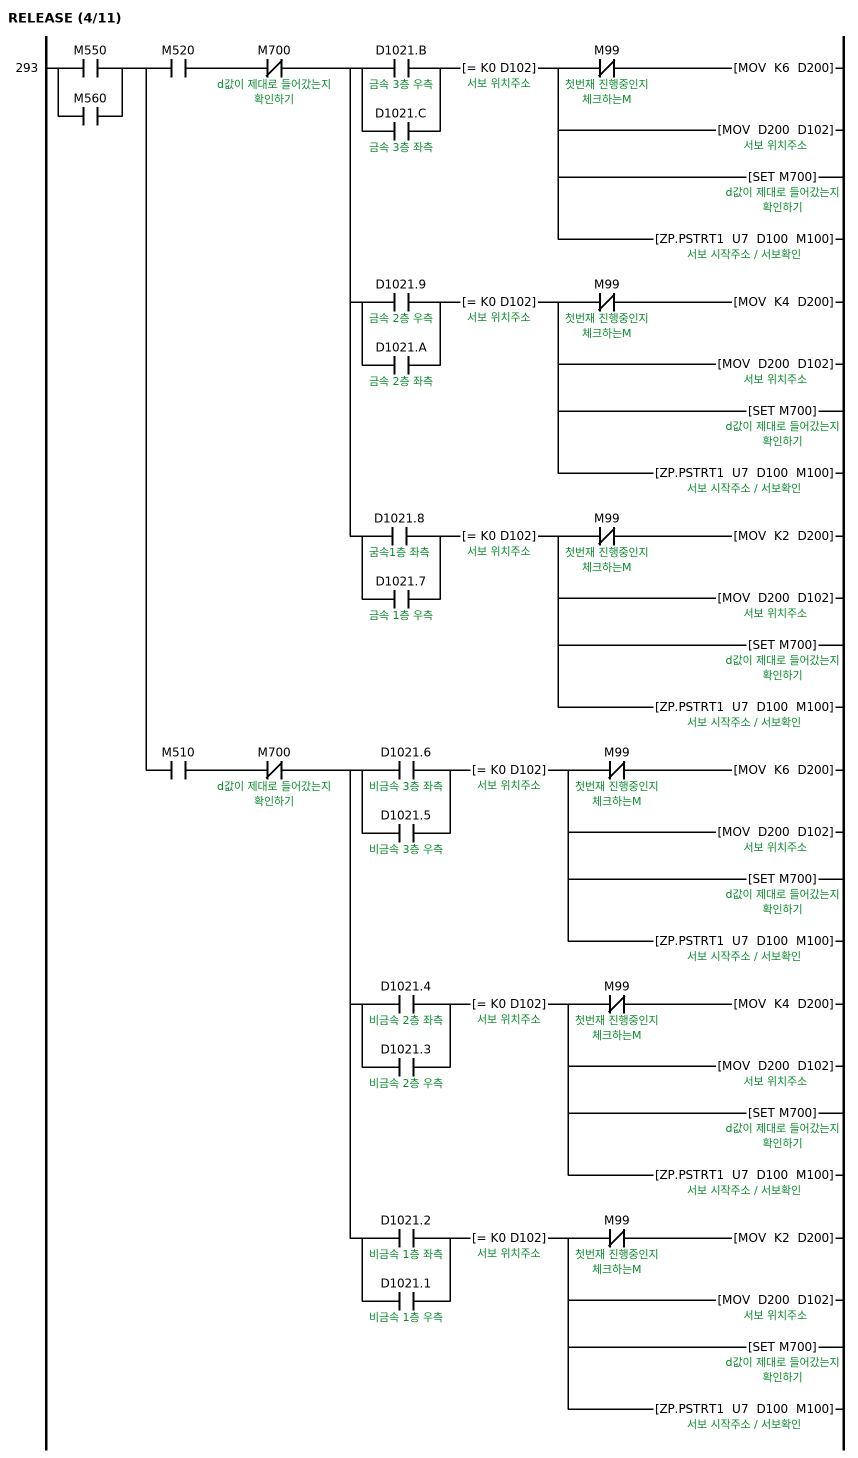
[picture p24: ladder of RELEASE, rungs at steps 293 to 293]
293   LD      M550
      OR      M560
      MPS
      AND     M520
      ANI     M700  ; d값이 제대로 들어갔는지 확인하기
      MPS
      LD      D1021.B  ; 금속 3층 우측
      OR      D1021.C  ; 금속 3층 좌측
      ANB
      AND=    K0 D102  ; 서보 위치주소
      MPS
      ANI     M99  ; 첫번재 진행중인지 체크하는M
      MOV     K6 D200
      MPP
      MOV     D200 D102
      SET     M700  ; d값이 제대로 들어갔는지 확인하기
      ZP.PSTRT1 U7 D100 M100  ; 서보 시작주소 / 서보확인
      MRD
      LD      D1021.9  ; 금속 2층 우측
      OR      D1021.A  ; 금속 2층 좌측
      ANB
      AND=    K0 D102  ; 서보 위치주소
      MPS
      ANI     M99  ; 첫번재 진행중인지 체크하는M
      MOV     K4 D200
      MPP
      MOV     D200 D102
      SET     M700  ; d값이 제대로 들어갔는지 확인하기
      ZP.PSTRT1 U7 D100 M100
      MPP
      LD      D1021.8  ; 굼속1층 좌측
      OR      D1021.7  ; 금속 1층 우측
      ANB
      AND=    K0 D102  ; 서보 위치주소
      MPS
      ANI     M99  ; 첫번재 진행중인지 체크하는M
      MOV     K2 D200
      MPP
      MOV     D200 D102
      SET     M700  ; d값이 제대로 들어갔는지 확인하기
      ZP.PSTRT1 U7 D100 M100
      MPP
      AND     M510
      ANI     M700  ; d값이 제대로 들어갔는지 확인하기
      MPS
      LD      D1021.6  ; 비금속 3층 좌측
      OR      D1021.5  ; 비금속 3층 우측
      ANB
      AND=    K0 D102  ; 서보 위치주소
      MPS
      ANI     M99  ; 첫번재 진행중인지 체크하는M
      MOV     K6 D200
      MPP
      MOV     D200 D102
      SET     M700  ; d값이 제대로 들어갔는지 확인하기
      ZP.PSTRT1 U7 D100 M100
      MRD
      LD      D1021.4  ; 비금속 2층 좌측
      OR      D1021.3  ; 비금속 2층 우측
      ANB
      AND=    K0 D102  ; 서보 위치주소
      MPS
      ANI     M99  ; 첫번재 진행중인지 체크하는M
      MOV     K4 D200
      MPP
      MOV     D200 D102
      SET     M700  ; d값이 제대로 들어갔는지 확인하기
      ZP.PSTRT1 U7 D100 M100
      MPP
      LD      D1021.2  ; 비금속 1층 좌측
      OR      D1021.1  ; 비금속 1층 우측
      ANB
      AND=    K0 D102  ; 서보 위치주소
      MPS
      ANI     M99  ; 첫번재 진행중인지 체크하는M
      MOV     K2 D200
      MPP
      MOV     D200 D102
      SET     M700  ; d값이 제대로 들어갔는지 확인하기
      ZP.PSTRT1 U7 D100 M100
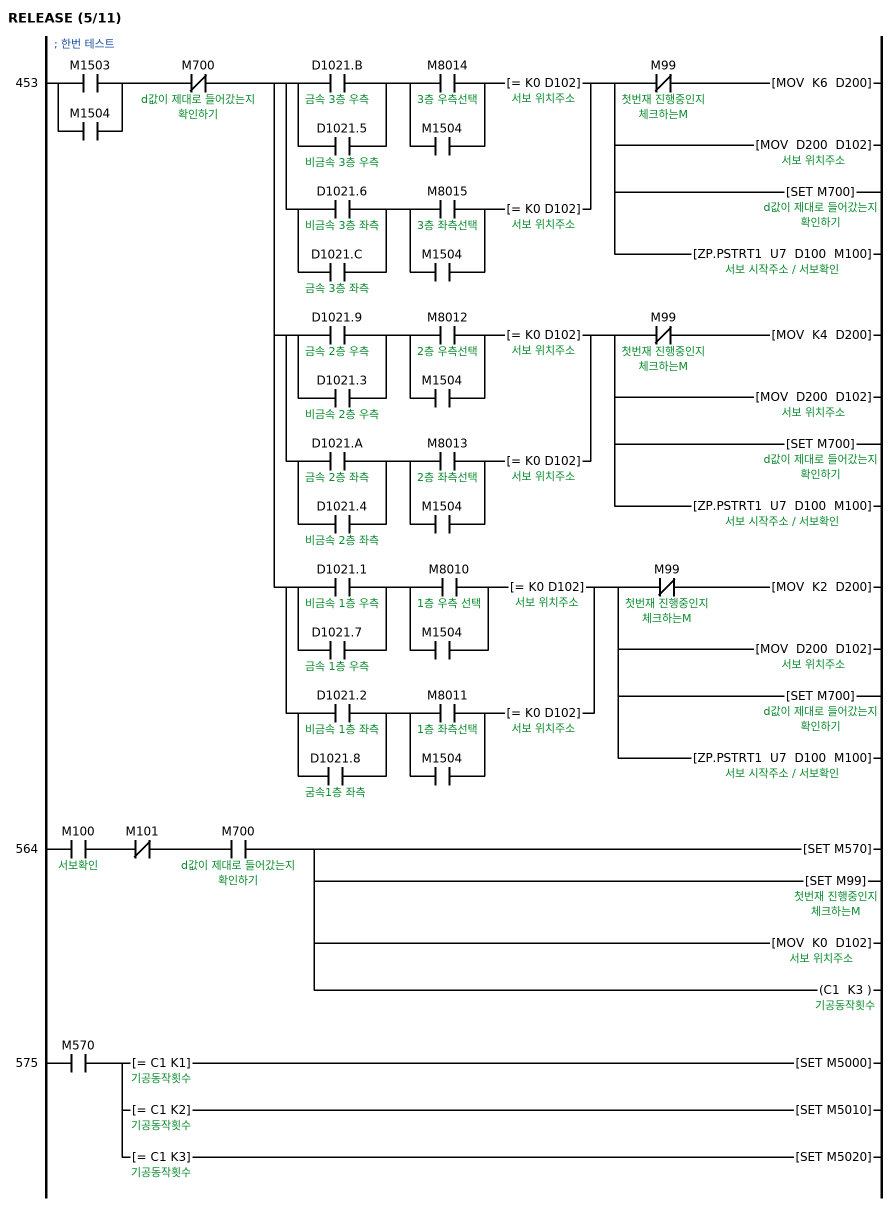
; 한번 테스트
453   LD      M1503
      OR      M1504
      ANI     M700  ; d값이 제대로 들어갔는지 확인하기
      MPS
      LD      D1021.B  ; 금속 3층 우측
      OR      D1021.5  ; 비금속 3층 우측
      LD      M8014  ; 3층 우측선택
      OR      M1504
      ANB
      AND=    K0 D102  ; 서보 위치주소
      LD      D1021.6  ; 비금속 3층 좌측
      OR      D1021.C  ; 금속 3층 좌측
      LD      M8015  ; 3층 좌측선택
      OR      M1504
      ANB
      AND=    K0 D102  ; 서보 위치주소
      ORB
      ANB
      MPS
      ANI     M99  ; 첫번재 진행중인지 체크하는M
      MOV     K6 D200
      MPP
      MOV     D200 D102
      SET     M700  ; d값이 제대로 들어갔는지 확인하기
      ZP.PSTRT1 U7 D100 M100
      MRD
      LD      D1021.9  ; 금속 2층 우측
      OR      D1021.3  ; 비금속 2층 우측
      LD      M8012  ; 2층 우측선택
      OR      M1504
      ANB
      AND=    K0 D102  ; 서보 위치주소
      LD      D1021.A  ; 금속 2층 좌측
      OR      D1021.4  ; 비금속 2층 좌측
      LD      M8013  ; 2층 좌측선택
      OR      M1504
      ANB
      AND=    K0 D102  ; 서보 위치주소
      ORB
      ANB
      MPS
      ANI     M99  ; 첫번재 진행중인지 체크하는M
      MOV     K4 D200
      MPP
      MOV     D200 D102
      SET     M700  ; d값이 제대로 들어갔는지 확인하기
      ZP.PSTRT1 U7 D100 M100
      MPP
      LD      D1021.1  ; 비금속 1층 우측
      OR      D1021.7  ; 금속 1층 우측
      LD      M8010  ; 1층 우측 선택
      OR      M1504
      ANB
      AND=    K0 D102  ; 서보 위치주소
      LD      D1021.2  ; 비금속 1층 좌측
      OR      D1021.8  ; 굼속1층 좌측
      LD      M8011  ; 1층 좌측선택
      OR      M1504
      ANB
      AND=    K0 D102  ; 서보 위치주소
      ORB
      ANB
      MPS
      ANI     M99  ; 첫번재 진행중인지 체크하는M
      MOV     K2 D200
      MPP
      MOV     D200 D102
      SET     M700  ; d값이 제대로 들어갔는지 확인하기
      ZP.PSTRT1 U7 D100 M100
564   LD      M100  ; 서보확인
      ANI     M101
      AND     M700  ; d값이 제대로 들어갔는지 확인하기
      SET     M570
      SET     M99  ; 첫번재 진행중인지 체크하는M
      MOV     K0 D102
      OUT     C1 K3  ; 기공동작횟수
575   LD      M570
      MPS
      AND=    C1 K1  ; 기공동작횟수
      SET     M5000
      MRD
      AND=    C1 K2  ; 기공동작횟수
      SET     M5010
      MPP
      AND=    C1 K3  ; 기공동작횟수
      SET     M5020
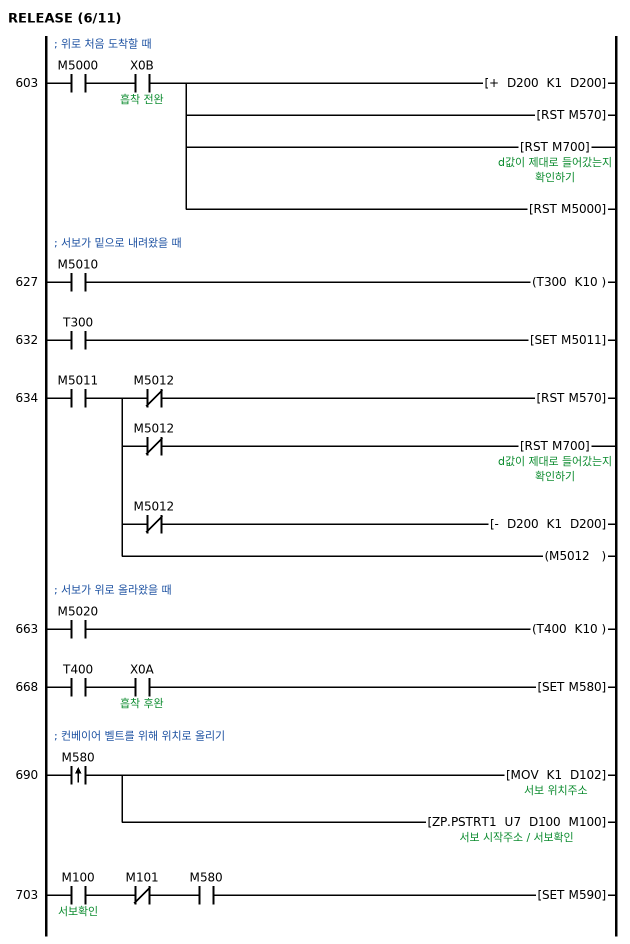
; 위로 처음 도착할 때
603   LD      M5000
      AND     X0B  ; 흡착 전완
      +       D200 K1 D200
      RST     M570
      RST     M700  ; d값이 제대로 들어갔는지 확인하기
      RST     M5000
; 서보가 밑으로 내려왔을 때
627   LD      M5010
      OUT     T300 K10
632   LD      T300
      SET     M5011
634   LD      M5011
      MPS
      ANI     M5012
      RST     M570
      MRD
      ANI     M5012
      RST     M700  ; d값이 제대로 들어갔는지 확인하기
      MRD
      ANI     M5012
      -       D200 K1 D200
      MPP
      OUT     M5012
; 서보가 위로 올라왔을 때
663   LD      M5020
      OUT     T400 K10
668   LD      T400
      AND     X0A  ; 흡착 후완
      SET     M580
; 컨베이어 벨트를 위해 위치로 올리기
690   LDP     M580
      MOV     K1 D102
      ZP.PSTRT1 U7 D100 M100
703   LD      M100  ; 서보확인
      ANI     M101
      AND     M580
      SET     M590
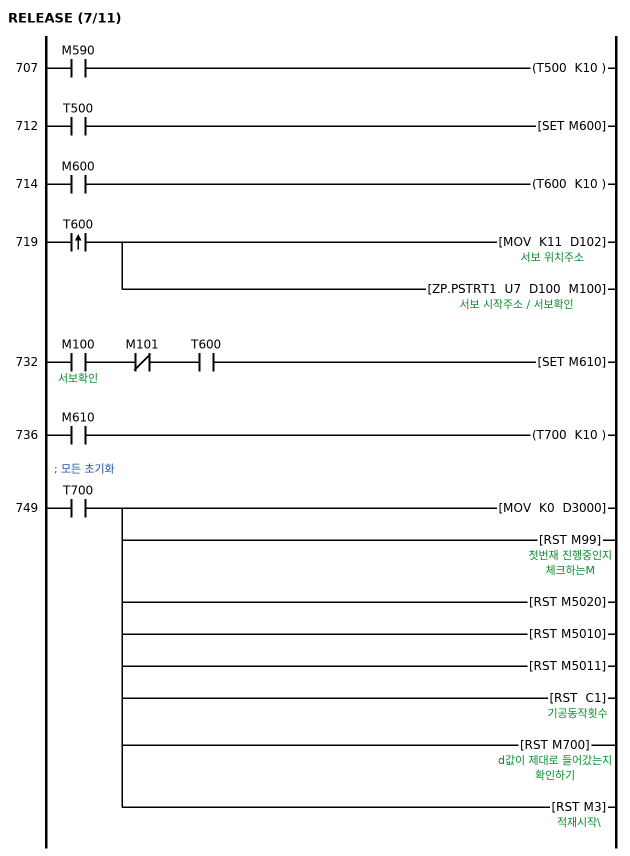
707   LD      M590
      OUT     T500 K10
712   LD      T500
      SET     M600
714   LD      M600
      OUT     T600 K10
719   LDP     T600
      MOV     K11 D102
      ZP.PSTRT1 U7 D100 M100
732   LD      M100  ; 서보확인
      ANI     M101
      AND     T600
      SET     M610
736   LD      M610
      OUT     T700 K10
; 모든 초기화
749   LD      T700
      MOV     K0 D3000
      RST     M99  ; 첫번재 진행중인지 체크하는M
      RST     M5020
      RST     M5010
      RST     M5011
      RST     C1  ; 기공동작횟수
      RST     M700  ; d값이 제대로 들어갔는지 확인하기
      RST     M3  ; 적재시작\
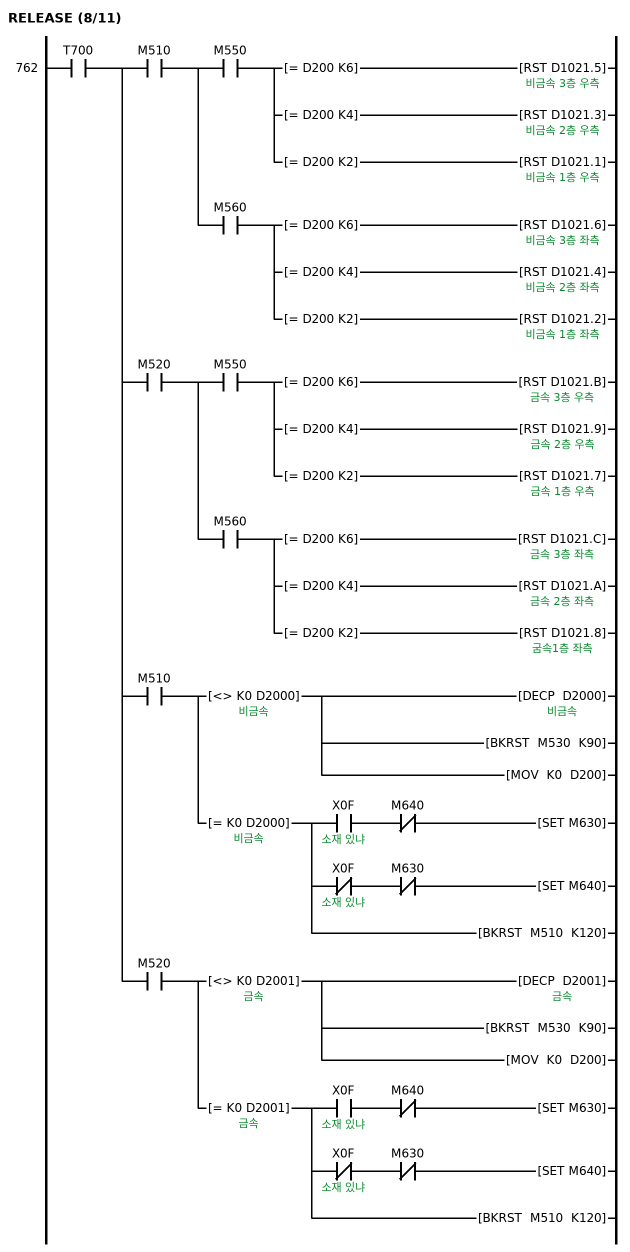
762   LD      T700
      MPS
      AND     M510
      MPS
      AND     M550
      MPS
      AND=    D200 K6
      RST     D1021.5  ; 비금속 3층 우측
      MRD
      AND=    D200 K4
      RST     D1021.3  ; 비금속 2층 우측
      MPP
      AND=    D200 K2
      RST     D1021.1  ; 비금속 1층 우측
      MPP
      AND     M560
      MPS
      AND=    D200 K6
      RST     D1021.6  ; 비금속 3층 좌측
      MRD
      AND=    D200 K4
      RST     D1021.4  ; 비금속 2층 좌측
      MPP
      AND=    D200 K2
      RST     D1021.2  ; 비금속 1층 좌측
      MRD
      AND     M520
      MPS
      AND     M550
      MPS
      AND=    D200 K6
      RST     D1021.B  ; 금속 3층 우측
      MRD
      AND=    D200 K4
      RST     D1021.9  ; 금속 2층 우측
      MPP
      AND=    D200 K2
      RST     D1021.7  ; 금속 1층 우측
      MPP
      AND     M560
      MPS
      AND=    D200 K6
      RST     D1021.C  ; 금속 3층 좌측
      MRD
      AND=    D200 K4
      RST     D1021.A  ; 금속 2층 좌측
      MPP
      AND=    D200 K2
      RST     D1021.8  ; 굼속1층 좌측
      MRD
      AND     M510
      MPS
      AND<>   K0 D2000  ; 비금속
      DECP    D2000
      BKRST   M530 K90
      MOV     K0 D200
      MPP
      AND=    K0 D2000  ; 비금속
      MPS
      AND     X0F  ; 소재 있냐
      ANI     M640
      SET     M630
      MRD
      ANI     X0F  ; 소재 있냐
      ANI     M630
      SET     M640
      MPP
      BKRST   M510 K120
      MPP
      AND     M520
      MPS
      AND<>   K0 D2001  ; 금속
      DECP    D2001
      BKRST   M530 K90
      MOV     K0 D200
      MPP
      AND=    K0 D2001  ; 금속
      MPS
      AND     X0F  ; 소재 있냐
      ANI     M640
      SET     M630
      MRD
      ANI     X0F  ; 소재 있냐
      ANI     M630
      SET     M640
      MPP
      BKRST   M510 K120
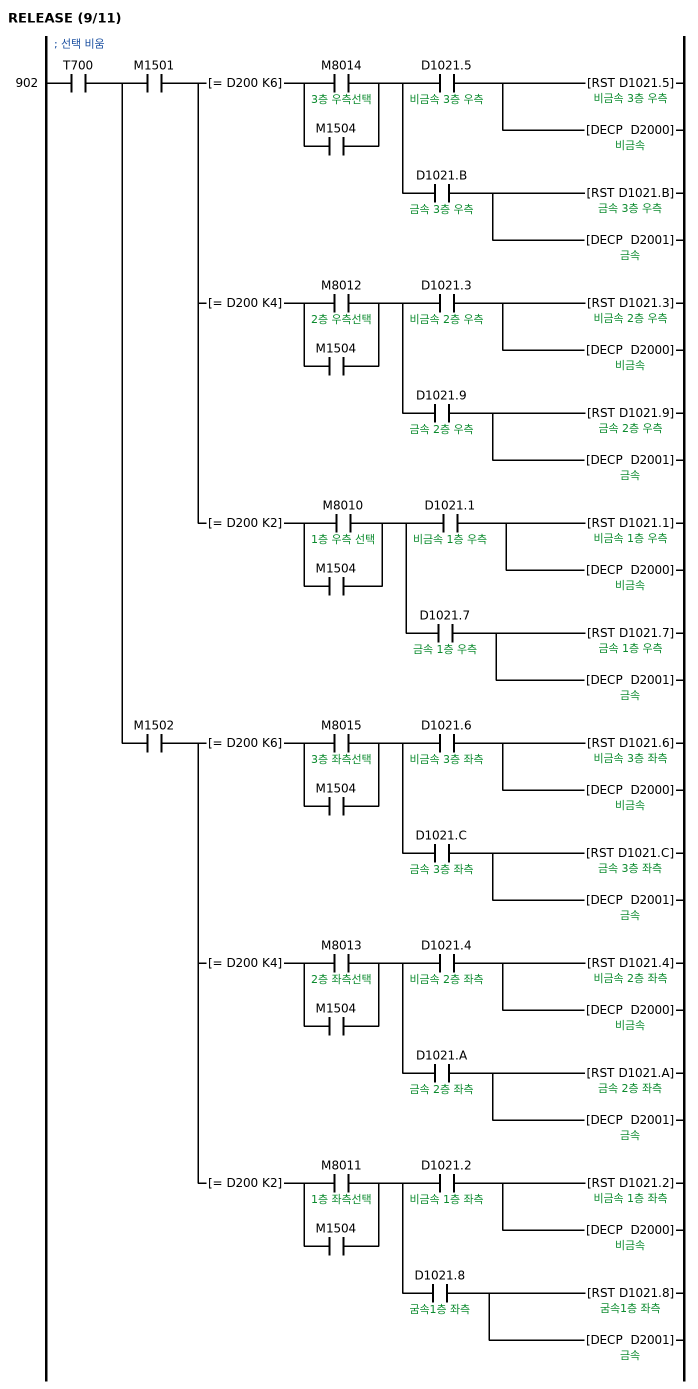
; 선택 비움
902   LD      T700
      MPS
      AND     M1501
      MPS
      AND=    D200 K6
      LD      M8014  ; 3층 우측선택
      OR      M1504
      ANB
      MPS
      AND     D1021.5  ; 비금속 3층 우측
      RST     D1021.5  ; 비금속 3층 우측
      DECP    D2000
      MPP
      AND     D1021.B  ; 금속 3층 우측
      RST     D1021.B  ; 금속 3층 우측
      DECP    D2001
      MRD
      AND=    D200 K4
      LD      M8012  ; 2층 우측선택
      OR      M1504
      ANB
      MPS
      AND     D1021.3  ; 비금속 2층 우측
      RST     D1021.3  ; 비금속 2층 우측
      DECP    D2000
      MPP
      AND     D1021.9  ; 금속 2층 우측
      RST     D1021.9  ; 금속 2층 우측
      DECP    D2001
      MPP
      AND=    D200 K2
      LD      M8010  ; 1층 우측 선택
      OR      M1504
      ANB
      MPS
      AND     D1021.1  ; 비금속 1층 우측
      RST     D1021.1  ; 비금속 1층 우측
      DECP    D2000
      MPP
      AND     D1021.7  ; 금속 1층 우측
      RST     D1021.7  ; 금속 1층 우측
      DECP    D2001
      MPP
      AND     M1502
      MPS
      AND=    D200 K6
      LD      M8015  ; 3층 좌측선택
      OR      M1504
      ANB
      MPS
      AND     D1021.6  ; 비금속 3층 좌측
      RST     D1021.6  ; 비금속 3층 좌측
      DECP    D2000
      MPP
      AND     D1021.C  ; 금속 3층 좌측
      RST     D1021.C  ; 금속 3층 좌측
      DECP    D2001
      MRD
      AND=    D200 K4
      LD      M8013  ; 2층 좌측선택
      OR      M1504
      ANB
      MPS
      AND     D1021.4  ; 비금속 2층 좌측
      RST     D1021.4  ; 비금속 2층 좌측
      DECP    D2000
      MPP
      AND     D1021.A  ; 금속 2층 좌측
      RST     D1021.A  ; 금속 2층 좌측
      DECP    D2001
      MPP
      AND=    D200 K2
      LD      M8011  ; 1층 좌측선택
      OR      M1504
      ANB
      MPS
      AND     D1021.2  ; 비금속 1층 좌측
      RST     D1021.2  ; 비금속 1층 좌측
      DECP    D2000
      MPP
      AND     D1021.8  ; 굼속1층 좌측
      RST     D1021.8  ; 굼속1층 좌측
      DECP    D2001
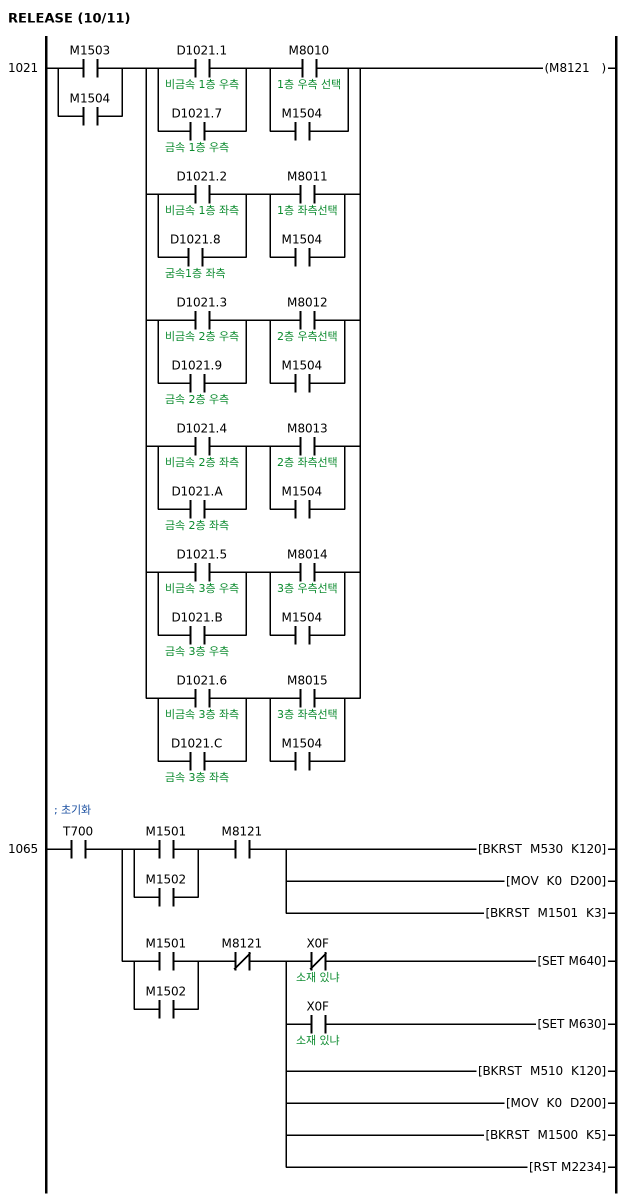
1021  LD      M1503
      OR      M1504
      LD      D1021.1  ; 비금속 1층 우측
      OR      D1021.7  ; 금속 1층 우측
      LD      M8010  ; 1층 우측 선택
      OR      M1504
      ANB
      LD      D1021.2  ; 비금속 1층 좌측
      OR      D1021.8  ; 굼속1층 좌측
      LD      M8011  ; 1층 좌측선택
      OR      M1504
      ANB
      ORB
      LD      D1021.3  ; 비금속 2층 우측
      OR      D1021.9  ; 금속 2층 우측
      LD      M8012  ; 2층 우측선택
      OR      M1504
      ANB
      ORB
      LD      D1021.4  ; 비금속 2층 좌측
      OR      D1021.A  ; 금속 2층 좌측
      LD      M8013  ; 2층 좌측선택
      OR      M1504
      ANB
      ORB
      LD      D1021.5  ; 비금속 3층 우측
      OR      D1021.B  ; 금속 3층 우측
      LD      M8014  ; 3층 우측선택
      OR      M1504
      ANB
      ORB
      LD      D1021.6  ; 비금속 3층 좌측
      OR      D1021.C  ; 금속 3층 좌측
      LD      M8015  ; 3층 좌측선택
      OR      M1504
      ANB
      ORB
      ANB
      OUT     M8121
; 초기화
1065  LD      T700
      MPS
      LD      M1501
      OR      M1502
      ANB
      AND     M8121
      BKRST   M530 K120
      MOV     K0 D200
      BKRST   M1501 K3
      MPP
      LD      M1501
      OR      M1502
      ANB
      ANI     M8121
      MPS
      ANI     X0F  ; 소재 있냐
      SET     M640
      MRD
      AND     X0F  ; 소재 있냐
      SET     M630
      MPP
      BKRST   M510 K120
      MOV     K0 D200
      BKRST   M1500 K5
      RST     M2234
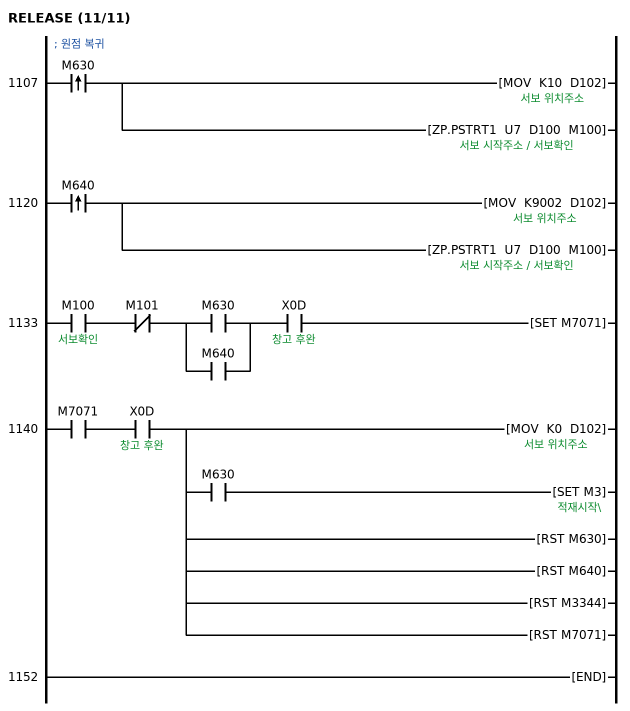
; 원점 복귀
1107  LDP     M630
      MOV     K10 D102
      ZP.PSTRT1 U7 D100 M100
1120  LDP     M640
      MOV     K9002 D102
      ZP.PSTRT1 U7 D100 M100
1133  LD      M100  ; 서보확인
      ANI     M101
      LD      M630
      OR      M640
      ANB
      AND     X0D  ; 창고 후완
      SET     M7071
1140  LD      M7071
      AND     X0D  ; 창고 후완
      MOV     K0 D102
      MPS
      AND     M630
      SET     M3  ; 적재시작\
      MPP
      RST     M630
      RST     M640
      RST     M3344
      RST     M7071
1152  END
END_PROGRAM

// device comments not shown above
X7  ; 배출 전완
X0C  ; 흡착 여부
X14  ; 컨베이어 엔코더 센서 감지
X16  ; Push Button2
X17  ; Push Button3
X18  ; Push Button4
X19  ; Push Button5
X1A  ; Push Button6
X1B  ; Push Button7
X1C  ; Toggle
Y25  ; 배출 전진
Y26  ; 배출 후진
M5  ; 비금 정리
M6  ; 적재시작
M10  ; 작업시작
M53  ; 창고 후진
M54  ; 창고 전진
M55  ; 창고 후진완료
M56  ; 창고 전진완료
M57  ; 카운트값 올려주는 M
M111  ; 비금속
M112  ; 금속
M200  ; 금속3우
M201  ; 금속3좌
M202  ; 금속2우
M203  ; 금속2좌
M204  ; 금속1우
M205  ; 금속1좌
M206  ; 비금3우
M207  ; 비금3좌
M208  ; 비금2우
M209  ; 비금2좌
M210  ; 비금1우
M211  ; 비금1좌
M710  ; 1층우버튼
M801  ; 3
M1023  ; HMI 수량초기화
M2223  ; 금속
M2224  ; 비금속
M4444  ; 실린더  초기상태X
M7676  ; 초기상태확인용
T1  ; 처음 실린더1초대기
T2  ; 비금속탐지 대기시간
T3  ; 서보 흡착 도착대기
T4  ; 위치상승후 대기
T5  ; 흡착 전진후 대기
T6  ; 컨베이어 시간
T7  ; 위치 상승후대기2
T10  ; 흡착대기시간
T11  ; 상승 대기 시간
T12  ; 흡착 전진후 대기시간
T13  ; 가공 대기
T14  ; 재상승 대기시잔
T15  ; 배출시간
T20  ; 비금속 컨베이어대기
T30  ; 배출
C2  ; 비금속 갯수
C3  ; 금속 갯수
D3  ; 목표위치
D1000  ; 목표위치
D1001  ; 현재위치
D1005  ; 현재 속도
D1009  ; 에러 번혼
D1010  ; 경고번호
D1011  ; 동작상태
D1020  ; 금속 수량
D1021  ; 비금속 수량
D1030  ; 가공 대기
D1031  ; 대기 시간
D1032  ; 가공 횟수
D1040  ; 가공 횟수
D5555  ; 램프 처리및 위치조절
D5556  ; 층수 처리
D5656  ; 금속 처리
D5657  ; 나머지
D5658  ; 비금속 처리
D5659  ; 비금속 나머지
D7011  ; 티칭 위치 인덱스
